TYPE E_TCPConnectionState :
(
	eTCP_STATE_IDLE,
	eTCP_STATE_CONNECT_START,
	eTCP_STATE_CONNECT_WAIT,
	eTCP_STATE_DATAEXCHANGE,
	eTCP_STATE_CLOSE_START,
	eTCP_STATE_CLOSE_WAIT,
	eTCP_STATE_ERROR
);
END_TYPE

(* stored: Version 1.1.0.1
   DUT E_TCPConnectionState: Id {ca07e5cf-6717-4474-a004-46cf1a6e254e} *)
